(* IEC 61131-3 sources: llm-plc-st-eval/data/processed_definitivo/gemini-3.1-pro-preview/I5/few_shot, 3 files *)

(* ---- ejec_1.st ---- *)
FUNCTION_BLOCK FB_Clasificadora
VAR_INPUT
    sensorPresencia : BOOL; (* Sensor de paso de pieza *)
    sensorAltura : BOOL;    (* Sensor de pieza alta *)
END_VAR
VAR_OUTPUT
    banda : BOOL;           (* Salida de la banda transportadora *)
    piston : BOOL;          (* Salida del piston desviador *)
    nAltas : INT;           (* Contador de piezas altas *)
    nBajas : INT;           (* Contador de piezas bajas *)
END_VAR
VAR
    trigPresencia : R_TRIG; (* Flanco de subida del sensor de presencia *)
    tpRetardo : TP;         (* Temporizador para el retardo de 2s *)
    ftrigRetardo : F_TRIG;  (* Flanco de bajada para detectar fin del retardo *)
    tpPiston : TP;          (* Temporizador para el pulso del piston de 1s *)
    piezaAlta : BOOL;       (* Marca temporal de pieza alta detectada *)
END_VAR

(* La banda funciona continuamente *)
banda := TRUE;

(* Deteccion de una nueva pieza (flanco de subida) *)
trigPresencia(CLK := sensorPresencia);

(* Clasificacion y conteo *)
piezaAlta := FALSE;
IF trigPresencia.Q THEN
    IF sensorAltura THEN
        nAltas := nAltas + 1;
        piezaAlta := TRUE; (* Dispara la secuencia del desviador *)
    ELSE
        nBajas := nBajas + 1;
    END_IF;
END_IF;

(* Retardo de 2 segundos al detectar una pieza alta *)
tpRetardo(IN := piezaAlta, PT := T#2S);

(* El fin del retardo genera un flanco de bajada *)
ftrigRetardo(CLK := tpRetardo.Q);

(* Pulso de 1 segundo para activar el piston desviador tras el retardo *)
tpPiston(IN := ftrigRetardo.Q, PT := T#1S);
piston := tpPiston.Q;

END_FUNCTION_BLOCK

(* ---- ejec_2.st ---- *)
FUNCTION_BLOCK FB_Clasificadora
VAR_INPUT
    sensorPresencia : BOOL; (* Detecta el paso de una pieza *)
    sensorAltura : BOOL;    (* Detecta si la pieza es alta *)
END_VAR
VAR_OUTPUT
    banda : BOOL;           (* Salida de la banda transportadora *)
    piston : BOOL;          (* Salida del piston desviador *)
    nAltas : INT;           (* Contador de piezas altas *)
    nBajas : INT;           (* Contador de piezas bajas *)
END_VAR
VAR
    flancoPresencia : R_TRIG; (* Detector de flanco para nueva pieza *)
    tpRetardo : TP;           (* Temporizador para el retardo de llegada (2s) *)
    finRetardo : F_TRIG;      (* Detector de fin del retardo *)
    tpPiston : TP;            (* Temporizador para la activacion del piston (1s) *)
    pulsoAlta : BOOL;         (* Marca interna para iniciar el retardo *)
END_VAR

(* La banda funciona continuamente *)
banda := TRUE;

(* Deteccion del paso de una nueva pieza *)
flancoPresencia(CLK := sensorPresencia);

pulsoAlta := FALSE;

(* Clasificacion y conteo al detectar la pieza *)
IF flancoPresencia.Q THEN
    IF sensorAltura THEN
        nAltas := nAltas + 1;
        pulsoAlta := TRUE; (* Inicia la secuencia de desvio *)
    ELSE
        nBajas := nBajas + 1;
    END_IF;
END_IF;

(* Genera un pulso de 2 segundos como retardo de llegada al desviador *)
tpRetardo(IN := pulsoAlta, PT := T#2S);

(* Detecta cuando terminan los 2 segundos de retardo *)
finRetardo(CLK := tpRetardo.Q);

(* Activa el piston durante 1 segundo justo al terminar el retardo *)
tpPiston(IN := finRetardo.Q, PT := T#1S);
piston := tpPiston.Q;

END_FUNCTION_BLOCK

(* ---- ejec_3.st ---- *)
FUNCTION_BLOCK FB_Clasificadora
VAR_INPUT
    sensorPresencia : BOOL; (* Sensor de paso de pieza *)
    sensorAltura : BOOL;    (* Sensor de pieza alta *)
END_VAR
VAR_OUTPUT
    banda : BOOL;           (* Salida de la banda transportadora *)
    piston : BOOL;          (* Salida del piston desviador *)
    nAltas : INT;           (* Contador de piezas altas *)
    nBajas : INT;           (* Contador de piezas bajas *)
END_VAR
VAR
    trigPresencia : R_TRIG; (* Flanco de subida del sensor de presencia *)
    pulsoAlta : BOOL;       (* Marca de deteccion de pieza alta *)
    tRetardo : TP;          (* Temporizador de retardo de llegada *)
    trigFinRetardo : F_TRIG;(* Flanco de bajada del retardo *)
    tPiston : TP;           (* Temporizador de activacion del piston *)
END_VAR

(* La banda funciona continuamente *)
banda := TRUE;

(* Detectar el paso de una nueva pieza *)
trigPresencia(CLK := sensorPresencia);

pulsoAlta := FALSE;
IF trigPresencia.Q THEN
    IF sensorAltura THEN
        nAltas := nAltas + 1;
        pulsoAlta := TRUE; (* Inicia la secuencia de desvio *)
    ELSE
        nBajas := nBajas + 1;
    END_IF;
END_IF;

(* Generar retardo de 2s desde la deteccion *)
tRetardo(IN := pulsoAlta, PT := T#2S);

(* Detectar el fin del retardo de 2s *)
trigFinRetardo(CLK := tRetardo.Q);

(* Activar el piston por 1s al terminar el retardo *)
tPiston(IN := trigFinRetardo.Q, PT := T#1S);
piston := tPiston.Q;

END_FUNCTION_BLOCK
